(*
SPDX-FileCopyrightText: © 2026 Oleksandr Tiutyk <trofimich@gmail.com>
SPDX-License-Identifier: MIT
License: https://opensource.org/license/mit
*)

(*!
<summary>Provides a resource-free task that counts one step per work call.</summary>
<description>
Configure the target before Start. A successful Reset from STOPPED clears the counter and retains the target.
</description>
*)

FUNCTION_BLOCK CounterTask EXTENDS TOF_Tasks.Task
VAR_STAT
	//! <summary>Class name shared by all instances of this function block.</summary>
	{attribute 'hide'} 
	_ClassName : STRING := __POUNAME();
END_VAR
VAR
	_Counter : INT;
	_TargetValue : INT;
END_VAR

{attribute 'monitoring' := 'call'}
PROPERTY ClassName : REFERENCE TO STRING
GET
ClassName REF= _ClassName;
END_GET
END_PROPERTY

{attribute 'monitoring' := 'call'}
PROPERTY Counter : INT
GET
Counter := _Counter;
END_GET
END_PROPERTY

{attribute 'monitoring' := 'call'}
PROPERTY NamespaceName : REFERENCE TO STRING
GET
NamespaceName REF= CurrentNamespace.Name;
END_GET
END_PROPERTY

METHOD PROTECTED OnRunning
VAR_OUTPUT
	processingState : TOF_Tasks.TASK_PROCESSING_STATE;
END_VAR
VAR_IN_OUT
	stopReasonMessage : TOF_Core.ERROR_MESSAGE;
END_VAR
_Counter := _Counter + 1;

IF _Counter >= _TargetValue THEN
	processingState := TOF_Tasks.TASK_PROCESSING_STATE.DONE;
END_IF
END_METHOD

(*!
<summary>Clears progress for a stopped counter while retaining its configured target.</summary>
<description>
Invoked by Task.Reset after termination. A counter prepared for the next run starts from zero.
</description>
*)
METHOD PROTECTED OnReset
_Counter := TOF_Core.SignedInt16.ZERO;
END_METHOD

{attribute 'monitoring' := 'call'}
PROPERTY SelfSize : ULINT
GET
SelfSize := XSIZEOF(THIS^);
END_GET
END_PROPERTY

{attribute 'monitoring' := 'call'}
PROPERTY TargetValue : INT
GET
TargetValue := _TargetValue;
END_GET
SET
_TargetValue := TargetValue;
END_SET
END_PROPERTY

END_FUNCTION_BLOCK

(* stored: Version 1.1.0.1, ProductVersion 3.1.4026.21
   POU CounterTask: Id {166c6948-6d4a-4978-a467-4fa58f366536}, SpecialFunc None
   Folder Overriden members: Id {97b0240c-e26a-4b1a-a761-8310302baa32}
   Property ClassName: Id {45e527f3-6e71-4c90-87c4-3da76042e202}
   Get Get: Id {877ce973-ecff-4501-891e-4e7fdafbe094}
   Property Counter: Id {346a7dae-aaf8-4179-a9b6-4ce063b5057f}
   Get Get: Id {b86ea06f-ce82-41b8-a812-d54bace1ff86}
   Property NamespaceName: Id {3229b47c-0917-45b8-af9a-5a06097fd17b}
   Get Get: Id {3db9af6e-af22-4f8b-afe9-58bd7358b5dd}
   Method OnRunning: Id {d8bd1379-eacd-49c3-be7f-5ac1efb7999d}
   Method OnReset: Id {6aa33ebe-c5ed-4315-9c11-cc7ec84291cf}
   Property SelfSize: Id {170d6f05-ca2a-424f-a507-a47e5aad4278}
   Get Get: Id {5cb9b1bb-9718-4868-bca8-98419f41a393}
   Property TargetValue: Id {acd773ca-12c6-4930-bbc0-7bd2cb5569b8}
   Get Get: Id {7d22ff02-01df-4b97-89d4-6f5f601f9b19}
   Set Set: Id {eca682e3-5906-4935-8b40-26af27e84e45} *)
